Staubli VAL3: utRectangle.dtx

public utBorder Border
  [0]
    string sBorderColour
    string sBorderWidth
public utAppearance Appearance
  [0]
    string sBackgroundColour
    string sColour
    bool bVisibility
public utCommon Common
  [0]
    bool bDisabled
    string sValue
    string sID
    num nValue
    string sPage
public utText Text
  [0]
    string sFontFamily
    string sFontStyle
    string sFontWeight
    string sTextAlignment
    num nFontSize
